{attribute 'qualified_only'}
{attribute 'strict'}
TYPE E_Piston_State :
(
	Init := 0,
	Close,Open,Busy_Close,Busy_Open
);
END_TYPE

(* stored: Version 1.1.0.1, ProductVersion 3.1.4024.12
   DUT E_Piston_State: Id {48fdafc9-fa88-4836-b7ef-d935a792ea8f} *)
